// TIA Portal V21 export
// export: Created 2026-11-10T22:39:24.158407Z, ExportSetting WithDefaults, DisplayName Totally Integrated Automation Portal, DisplayVersion V21 Update 3, DisplayName STEP 7 Professional, DisplayVersion V21 Update 3, DisplayName STEP 7 Safety, DisplayVersion V21, DisplayName Tech WebApplication, DisplayVersion V21, DisplayName WinCC Basic/Comfort/Advanced, DisplayVersion V21 Update 3, DisplayName WinCC Unified, DisplayVersion V21 Update 3
DATA_BLOCK "mTO_SynchronousAxis"   // DB8, Motion_DB
// stored: AutoNumber true, DBAccessibleFromOPCUA true, DBAccessibleFromWebserver true, InstanceOfName TO_SynchronousAxis_2, OfSystemLibElement TO_SynchronousAxis, OfSystemLibVersion 6.0
TO_SynchronousAxis_2   // technology object, version 6.0
// stored: Connection Interface Actor
// stored: Connection Interface Sensor[1]
// stored: Connection Interface Torque
   // // inherited from TO_PositioningAxis
   // // inherited from TO_SpeedAxis
   // // inherited from TO_Axis
   // // inherited from TO_Object
   // VAR
   //    Velocity : LReal;
   //    Acceleration : LReal;
   //    ActualSpeed : LReal;
   //    VelocitySetpoint : LReal;
   //    Actor : TO_Struct_Actor;
   //    TorqueLimiting : TO_Struct_TorqueLimiting;
   //    LoadGear : TO_Struct_LoadGear;
   //    DynamicLimits : TO_Struct_DynamicLimits;
   //    DynamicDefaults : TO_Struct_DynamicDefaults;
   //    Override : TO_Struct_Override;
   //    Units : TO_Struct_Units;
   //    StatusDrive : TO_Struct_StatusDrive;
   //    StatusTorqueData : TO_Struct_StatusTorqueData;
   //    StatusMotionIn : TO_Struct_StatusMotionIn;
   //    StatusWord : DWord;
   //    StatusWord2 : DWord;
   //    ErrorWord : DWord;
   //    ErrorDetail : TO_Struct_ErrorDetail;
   //    WarningWord : DWord;
   //    ControlPanel : TO_Struct_ControlPanel;
   //    InternalToTrace : Array[1..4] of TO_Struct_Internal;
   //    VirtualAxis : TO_Struct_VirtualAxis;
   //    Simulation : TO_Struct_AxisSimulation;
   // END_VAR
   // VAR
   //    Position : LReal;
   //    ActualPosition : LReal;
   //    ActualVelocity : LReal;
   //    ActualAcceleration : LReal;
   //    OperativeSensor : UDInt;
   //    ModuloCycle : DInt;
   //    ActualModuloCycle : DInt;
   //    Clamping : TO_Struct_Clamping;
   //    Sensor : Array[1..4] of TO_Struct_Sensor;
   //    Extrapolation : TO_Struct_Extrapolation;
   //    Mechanics : TO_Struct_Mechanics;
   //    Properties : TO_Struct_Properties;
   //    Modulo : TO_Struct_Modulo;
   //    PositionLimits_SW : TO_Struct_PositionLimitsSW;
   //    PositionLimits_HW : TO_Struct_PositionLimitsHW;
   //    Homing : TO_Struct_Homing;
   //    PositionControl : TO_Struct_PositionControl;
   //    DynamicAxisModel : TO_Struct_DynamicAxisModel;
   //    FollowingError : TO_Struct_FollowingError;
   //    CrossPlcSynchronousOperation : TO_Struct_CrossPlcSynchronousOperation;
   //    PositioningMonitoring : TO_Struct_PositioningMonitoring;
   //    StandstillSignal : TO_Struct_StandstillSignal;
   //    StatusPositioning : TO_Struct_StatusPositioning;
   //    StatusServo : TO_Struct_StatusServo;
   //    StatusProvidedLeadingValue : TO_Struct_StatusProvidedLeadingValue;
   //    StatusSensor : Array[1..4] of TO_Struct_StatusSensor;
   //    StatusExtrapolation : TO_Struct_StatusExtrapolation;
   //    StatusKinematicsMotion : TO_Struct_StatusKinematicsMotion;
   // END_VAR
   // VAR
   //    StatusSynchronizedMotion { ExternalWritable := 'False'; S7_SetPoint := 'True'} : TO_Struct_StatusSynchronizedMotion;
   // END_VAR
BEGIN
   VirtualAxis.Mode := 1;
   VirtualAxis.Mode := 1;
END_DATA_BLOCK
